// TIA Portal V20 export
// export: Created 2026-11-12T11:17:34.1179187Z, ExportSetting WithDefaults, DisplayName Totally Integrated Automation Portal, DisplayVersion V20, DisplayName TIA Portal Openness, DisplayVersion V20, DisplayName TIA Portal Teamcenter Gateway, DisplayVersion V20, DisplayName TIA Portal Version Control Interface, DisplayVersion V20, DisplayName STEP 7 Professional, DisplayVersion V20, DisplayName STEP 7 CFC, DisplayVersion V20, DisplayName STEP 7 Safety, DisplayVersion V20, DisplayName WinCC Basic/Comfort/Advanced, DisplayVersion V20, DisplayName SIMATIC Visualization Architect, DisplayVersion V20, DisplayName WinCC Professional, DisplayVersion V20, DisplayName SIMATIC Visualization Architect, DisplayVersion V20, DisplayName WinCC Unified, DisplayVersion V20, DisplayName SIMATIC Visualization Architect, DisplayVersion V20
TYPE "UDT_Salidas_Basico"
// stored: IsFailsafeCompliant false
   STRUCT
      Led_boton_marcha : Bool;   // Luz del boton de Marcha
      Led_boton_rearme : Bool;   // Luz del boton de Reset
      Led_q1_ciclo_auto : Bool;   // Luz Q1
      Led_q2_emergencia : Bool;   // Luz Q2
      Cinta_dch : Bool;   // Arrancar cinta hacia la derecha
      Cinta_izq : Bool;   // Arrancar cinta hacia la izquierda
      Cinta_velocidad_baja : Bool;   // Establecer velocidad baja
      Bajar_stopper : Bool;   // Bajar cilindro Stopper
   END_STRUCT;
END_TYPE
